TYPE "ST_ModePolicy"
VERSION : 0.1
   STRUCT
      Shield : DInt;
      Style : DInt;
   END_STRUCT;

END_TYPE

